// TIA Portal V21 export
DATA_BLOCK "IDB_AnaDoubleAssign"   // DB10
// stored: InstanceOfName FB_AnaDoubleAssign, InstanceOfType FB
"FB_AnaDoubleAssign"
   // VAR_INPUT
   //    Start : Bool;
   //    Stop : Bool;
   // END_VAR
   // VAR_OUTPUT
   //    Motor : Bool;
   // END_VAR
BEGIN
END_DATA_BLOCK
